(* IEC 61131-3 sources: POMIRTS_lab3/AS/Library_2/ArCert, 3 files *)

(* ---- ArCert.typ ---- *)
 TYPE
	ArCertDetailsType : STRUCT				(*certificate details*)
		Name			: STRING[255]; 			(*certificate name*)
		Issuer			: STRING[255];			(*issuer (CN)*)
		Subject			: STRING[255];			(*subject (CN)*)
		ValidFrom		: DTStructure;			(*valid from date*)
		ValidTo			: DTStructure;			(*valid to date*)
		Version			: DINT;					(*version*)
		SerialNumber	: STRING[39];			(*serial number*)
	END_STRUCT;

	ArCertCRLDetailsType : STRUCT			(*detail information of a certificate revocation list (CRL)*)
		Name			: STRING[255]; 			(*CRL name*)
		Issuer			: STRING[255]; 			(*issuer*)
		EffectiveDate	: DTStructure;			(*effective date*)
		NextUpdate		: DTStructure;			(*next update*)
		Version			: DINT;					(*version*)
		CRLNumber      	: STRING[39]; 			(*CRL number*)
	END_STRUCT;

    ArCertKeySizeEnum :
        (
            arCERT_KEY_SIZE_1024_BITS := 1,		(*encryption with a key with 1024 bits*)
            arCERT_KEY_SIZE_2048_BITS := 2,		(*encryption with a key with 2048 bits*)
            arCERT_KEY_SIZE_4096_BITS := 3		(*encryption with a key with 4096 bits*)
        );

    ArCertAsyncInternalType : STRUCT
        FBStateCtx		: ArFBStateInternalType;
		AsyFuMaCtx		: ArFBAsyFuMaInternalType;
    END_STRUCT;
END_TYPE

(* ---- ArCert.fun ---- *)
{REDUND_CONTEXT} {REDUND_UNREPLICABLE} FUNCTION_BLOCK ArCertImportOwn   				(*imports an existing own certificate from buffer*)
	VAR_INPUT
		Execute			: BOOL; 			(*starts execution*) 			(**) (*#PAR*)
		Name 			: STRING[255];		(*name of the own certificate*) 	(**) (*#PAR*)
		Data			: UDINT; 			(*pointer to certificate data*) (**) (*#PAR*)
		DataSize 		: UDINT;			(*size of certificate data*) 	(**) (*#PAR*)
	END_VAR
	VAR_OUTPUT
		Done			: BOOL;				(*execution done*) 				(**) (*#PAR*)
		Busy			: BOOL;				(*execution running*) 			(**) (*#PAR*)
		Error			: BOOL;				(*execution failed*) 			(**) (*#PAR*)
		StatusID		: DINT;  			(*execution error: see help*) 	(**) (*#PAR*)
	END_VAR
	VAR
		Internal		: ArCertAsyncInternalType;	(*internal variable*)
	END_VAR
END_FUNCTION_BLOCK

{REDUND_CONTEXT} {REDUND_UNREPLICABLE} FUNCTION_BLOCK ArCertExportOwn  				(*exports an own certificate to a buffer*)
	VAR_INPUT
		Execute			: BOOL; 			(*starts execution*) 			(**) (*#PAR*)
		Name 			: STRING[255];		(*name of the own certificate*) 	(**) (*#PAR*)
		Data			: UDINT; 			(*pointer to buffer for exported certificate data*) (**) (*#PAR*)
		DataSize		: UDINT;			(*buffer size*) 				(**) (*#PAR*)
	END_VAR
	VAR_OUTPUT
		Done			: BOOL;				(*execution done*) 				(**) (*#PAR*)
		Busy			: BOOL;				(*execution running*) 			(**) (*#PAR*)
		Error			: BOOL;				(*execution failed*) 			(**) (*#PAR*)
		StatusID		: DINT;  			(*execution error: see help*) 	(**) (*#PAR*)
		NeededDataSize 	: UDINT;			(*needed buffer size*) 				(**) (*#PAR*)
	END_VAR
	VAR
		Internal		: ArCertAsyncInternalType;	(*internal variable*)
	END_VAR
END_FUNCTION_BLOCK

{REDUND_CONTEXT} {REDUND_UNREPLICABLE} FUNCTION_BLOCK ArCertDeleteOwn  				(*deletes an own certificate*)
	VAR_INPUT
		Execute			: BOOL; 			(*starts execution*) 			(**) (*#PAR*)
		Name 			: STRING[255];		(*name of the own certificate*) 	(**) (*#PAR*)
	END_VAR
	VAR_OUTPUT
		Done			: BOOL;				(*execution done*) 				(**) (*#PAR*)
		Busy			: BOOL;				(*execution running*) 			(**) (*#PAR*)
		Error			: BOOL;				(*execution failed*) 			(**) (*#PAR*)
		StatusID		: DINT;  			(*execution error: see help*) 	(**) (*#PAR*)
	END_VAR
	VAR
		Internal		: ArCertAsyncInternalType;	(*internal variable*)
	END_VAR
END_FUNCTION_BLOCK

{REDUND_CONTEXT} {REDUND_UNREPLICABLE} FUNCTION_BLOCK ArCertImportThirdParty   				(*imports an existing third party certificate from buffer*)
	VAR_INPUT
		Execute			: BOOL; 			(*starts execution*) 			(**) (*#PAR*)
		Name 			: STRING[255];		(*name of the third party certificate*) 	(**) (*#PAR*)
		Data			: UDINT; 			(*pointer to certificate data*) (**) (*#PAR*)
		DataSize 		: UDINT;			(*size of certificate data*) 	(**) (*#PAR*)
	END_VAR
	VAR_OUTPUT
		Done			: BOOL;				(*execution done*) 				(**) (*#PAR*)
		Busy			: BOOL;				(*execution running*) 			(**) (*#PAR*)
		Error			: BOOL;				(*execution failed*) 			(**) (*#PAR*)
		StatusID		: DINT;  			(*execution error: see help*) 	(**) (*#PAR*)
	END_VAR
	VAR
		Internal		: ArCertAsyncInternalType;	(*internal variable*)
	END_VAR
END_FUNCTION_BLOCK

{REDUND_CONTEXT} {REDUND_UNREPLICABLE} FUNCTION_BLOCK ArCertExportThirdParty  				(*exports a third party certificate to a buffer*)
	VAR_INPUT
		Execute			: BOOL; 			(*starts execution*) 			(**) (*#PAR*)
		Name 			: STRING[255];		(*name of the third party certificate*) 	(**) (*#PAR*)
		Data			: UDINT; 			(*pointer to buffer for exported certificate data*) (**) (*#PAR*)
		DataSize		: UDINT;			(*buffer size*) 				(**) (*#PAR*)
	END_VAR
	VAR_OUTPUT
		Done			: BOOL;				(*execution done*) 				(**) (*#PAR*)
		Busy			: BOOL;				(*execution running*) 			(**) (*#PAR*)
		Error			: BOOL;				(*execution failed*) 			(**) (*#PAR*)
		StatusID		: DINT;  			(*execution error: see help*) 	(**) (*#PAR*)
		NeededDataSize 	: UDINT;			(*needed buffer size*) 				(**) (*#PAR*)
	END_VAR
	VAR
		Internal		: ArCertAsyncInternalType;	(*internal variable*)
	END_VAR
END_FUNCTION_BLOCK

{REDUND_CONTEXT} {REDUND_UNREPLICABLE} FUNCTION_BLOCK ArCertDeleteThirdParty  				(*deletes a third party certificate*)
	VAR_INPUT
		Execute			: BOOL; 			(*starts execution*) 			(**) (*#PAR*)
		Name 			: STRING[255];		(*name of the third party certificate*) 	(**) (*#PAR*)
	END_VAR
	VAR_OUTPUT
		Done			: BOOL;				(*execution done*) 				(**) (*#PAR*)
		Busy			: BOOL;				(*execution running*) 			(**) (*#PAR*)
		Error			: BOOL;				(*execution failed*) 			(**) (*#PAR*)
		StatusID		: DINT;  			(*execution error: see help*) 	(**) (*#PAR*)
	END_VAR
	VAR
		Internal		: ArCertAsyncInternalType;	(*internal variable*)
	END_VAR
END_FUNCTION_BLOCK

{REDUND_CONTEXT} {REDUND_UNREPLICABLE} FUNCTION_BLOCK ArCertImportPrivateKey		(*imports an existing private key from buffer*)
	VAR_INPUT
		Execute			: BOOL; 			(*starts execution*) 			(**) (*#PAR*)
		Name 			: STRING[255];		(*name of the private key*) 	(**) (*#PAR*)
		Data			: UDINT; 			(*pointer to private key data*) (**) (*#PAR*)
		DataSize 		: UDINT;			(*size of private key data*) 	(**) (*#PAR*)
	END_VAR
	VAR_OUTPUT
		Done			: BOOL;				(*execution done*) 				(**) (*#PAR*)
		Busy			: BOOL;				(*execution running*) 			(**) (*#PAR*)
		Error			: BOOL;				(*execution failed*) 			(**) (*#PAR*)
		StatusID		: DINT;  			(*execution error: see help*) 	(**) (*#PAR*)
	END_VAR
	VAR
		Internal		: ArCertAsyncInternalType;	(*internal variable*)
	END_VAR
END_FUNCTION_BLOCK

{REDUND_CONTEXT} {REDUND_UNREPLICABLE} FUNCTION_BLOCK ArCertExportPrivateKey  		(*exports a private key to a buffer*)
	VAR_INPUT
		Execute			: BOOL; 			(*starts execution*) 			(**) (*#PAR*)
		Name 			: STRING[255];		(*name of the private key*) 	(**) (*#PAR*)
		Data			: UDINT; 			(*pointer to buffer for exported private key data*) (**) (*#PAR*)
		DataSize		: UDINT;			(*buffer size*) 				(**) (*#PAR*)
	END_VAR
	VAR_OUTPUT
		Done			: BOOL;				(*execution done*) 				(**) (*#PAR*)
		Busy			: BOOL;				(*execution running*) 			(**) (*#PAR*)
		Error			: BOOL;				(*execution failed*) 			(**) (*#PAR*)
		StatusID		: DINT;  			(*execution error: see help*) 	(**) (*#PAR*)
		NeededDataSize 	: UDINT;			(*needed buffer size*) 				(**) (*#PAR*)
	END_VAR
	VAR
		Internal		: ArCertAsyncInternalType;	(*internal variable*)
	END_VAR
END_FUNCTION_BLOCK

{REDUND_CONTEXT} {REDUND_UNREPLICABLE} FUNCTION_BLOCK ArCertDeletePrivateKey		(*deletes a private key*)
	VAR_INPUT
		Execute			: BOOL; 			(*starts execution*) 			(**) (*#PAR*)
		Name 			: STRING[255];		(*name of the private key*) 	(**) (*#PAR*)
	END_VAR
	VAR_OUTPUT
		Done			: BOOL;				(*execution done*) 				(**) (*#PAR*)
		Busy			: BOOL;				(*execution running*) 			(**) (*#PAR*)
		Error			: BOOL;				(*execution failed*) 			(**) (*#PAR*)
		StatusID		: DINT;  			(*execution error: see help*) 	(**) (*#PAR*)
	END_VAR
	VAR
		Internal		: ArCertAsyncInternalType;	(*internal variable*)
	END_VAR
END_FUNCTION_BLOCK

{REDUND_CONTEXT} {REDUND_UNREPLICABLE} FUNCTION_BLOCK ArCertImportCRL 				(*imports a certificate revocation list from buffer*)
	VAR_INPUT
		Execute			: BOOL; 			(*starts execution*) 			(**) (*#PAR*)
		Name 			: STRING[255];		(*name of the certificate revocation list*) 	(**) (*#PAR*)
		Data			: UDINT; 			(*pointer to certificate data*) (**) (*#PAR*)
		DataSize 		: UDINT;			(*size of certificate data*) 	(**) (*#PAR*)
	END_VAR
	VAR_OUTPUT
		Done			: BOOL;				(*execution done*) 				(**) (*#PAR*)
		Busy			: BOOL;				(*execution running*) 			(**) (*#PAR*)
		Error			: BOOL;				(*execution failed*) 			(**) (*#PAR*)
		StatusID		: DINT;  			(*execution error: see help*) 	(**) (*#PAR*)
	END_VAR
	VAR
		Internal		: ArCertAsyncInternalType;	(*internal variable*)
	END_VAR
END_FUNCTION_BLOCK

{REDUND_CONTEXT} {REDUND_UNREPLICABLE} FUNCTION_BLOCK ArCertExportCRL 				(*exports a certificate revocation list to a buffer*)
	VAR_INPUT
		Execute			: BOOL; 			(*starts execution*) 			(**) (*#PAR*)
		Name 			: STRING[255];		(*name of the certificate revocation list*) 	(**) (*#PAR*)
		Data			: UDINT; 			(*pointer to buffer for exported CRL data*) (**) (*#PAR*)
		DataSize		: UDINT;			(*buffer size*) 				(**) (*#PAR*)
	END_VAR
	VAR_OUTPUT
		Done			: BOOL;				(*execution done*) 				(**) (*#PAR*)
		Busy			: BOOL;				(*execution running*) 			(**) (*#PAR*)
		Error			: BOOL;				(*execution failed*) 			(**) (*#PAR*)
		StatusID		: DINT;  			(*execution error: see help*) 	(**) (*#PAR*)
		NeededDataSize : UDINT;				(*needed buffer size*) 				(**) (*#PAR*)
	END_VAR
	VAR
		Internal		: ArCertAsyncInternalType;	(*internal variable*)
	END_VAR
END_FUNCTION_BLOCK

{REDUND_CONTEXT} {REDUND_UNREPLICABLE} FUNCTION_BLOCK ArCertDeleteCRL  			(*deletes a certificate revocation list*)
	VAR_INPUT
		Execute			: BOOL; 			(*starts execution*) 			(**) (*#PAR*)
		Name 			: STRING[255];		(*name of the certificate revocation list*) 	(**) (*#PAR*)
	END_VAR
	VAR_OUTPUT
		Done			: BOOL;				(*execution done*) 				(**) (*#PAR*)
		Busy			: BOOL;				(*execution running*) 			(**) (*#PAR*)
		Error			: BOOL;				(*execution failed*) 			(**) (*#PAR*)
		StatusID		: DINT;  			(*execution error: see help*) 	(**) (*#PAR*)
	END_VAR
	VAR
		Internal		: ArCertAsyncInternalType;	(*internal variable*)
	END_VAR
END_FUNCTION_BLOCK

{REDUND_CONTEXT} {REDUND_UNREPLICABLE} FUNCTION_BLOCK ArCertGenerate       		(*generates a self-signed certificate and a private key*)
	VAR_INPUT
		Execute			: BOOL; 			(*starts execution*) 			(**) (*#PAR*)
		Name 			: STRING[255];		(*name of the certificate*) 	(**) (*#PAR*)
		PrivateKeyName 	: STRING[255];		(*name of the private key*) 	(**) (*#PAR*)
		KeySize 		: ArCertKeySizeEnum;(*size of key for certificate generation*) 	(**) (*#PAR*)
		CountryCode		: STRING[9];		(*country code*)		 		(**) (*#PAR*)
		StateProvince	: STRING[513];		(*state*) 						(**) (*#PAR*)
		Locality		: STRING[513];		(*locality*) 					(**) (*#PAR*)
		Organization 	: STRING[255];		(*organization*) 				(**) (*#PAR*)
		OrganizationUnit: STRING[255];		(*organization unit*) 			(**) (*#PAR*)
		ContactEmail 	: STRING[513];		(*contact email*)			 	(**) (*#PAR*)
		CommonName 		: STRING[255];		(*common name*) 				(**) (*#PAR*)
		ValidTimeSeconds : UDINT;			(*valid time in seconds*)		(**) (*#PAR*)
	END_VAR
	VAR_OUTPUT
		Done			: BOOL;				(*execution done*) 				(**) (*#PAR*)
		Busy			: BOOL;				(*execution running*) 			(**) (*#PAR*)
		Error			: BOOL;				(*execution failed*) 			(**) (*#PAR*)
		StatusID		: DINT;  			(*execution error: see help*) 	(**) (*#PAR*)
	END_VAR
	VAR
		Internal		: ArCertAsyncInternalType;	(*internal variable*)
	END_VAR
END_FUNCTION_BLOCK

{REDUND_CONTEXT} {REDUND_UNREPLICABLE} FUNCTION_BLOCK ArCertGenerateOpcUA		(*generates a self-signed certificate and a private key*)
	VAR_INPUT
		Execute			: BOOL; 			(*starts execution*) 			(**) (*#PAR*)
		Name 			: STRING[255];		(*name of the certificate*) 	(**) (*#PAR*)
		PrivateKeyName 	: STRING[255];		(*name of the private key*) 	(**) (*#PAR*)
		PrivateKeyPassword : STRING[255];	(*password of the private key*) (**) (*#PAR*)
		KeySize 		: ArCertKeySizeEnum;(*size of key for certificate generation*) 	(**) (*#PAR*)
		CountryCode		: STRING[9];		(*country code*)		 		(**) (*#PAR*)
		StateProvince	: STRING[513];		(*state*) 						(**) (*#PAR*)
		Locality		: STRING[513];		(*locality*) 					(**) (*#PAR*)
		Organization 	: STRING[255];		(*organization*) 				(**) (*#PAR*)
		OrganizationUnit: STRING[255];		(*organization unit*) 			(**) (*#PAR*)
		ContactEmail 	: STRING[513];		(*contact email*)			 	(**) (*#PAR*)
		CommonName 		: STRING[255];		(*common name*) 				(**) (*#PAR*)
		ValidTimeSeconds : UDINT;			(*valid time in seconds*)		(**) (*#PAR*)
		URI				: STRING[255];		(*URI*) 						(**) (*#PAR*)
	END_VAR
	VAR_OUTPUT
		Done			: BOOL;				(*execution done*) 				(**) (*#PAR*)
		Busy			: BOOL;				(*execution running*) 			(**) (*#PAR*)
		Error			: BOOL;				(*execution failed*) 			(**) (*#PAR*)
		StatusID		: DINT;  			(*execution error: see help*) 	(**) (*#PAR*)
	END_VAR
	VAR
		Internal		: ArCertAsyncInternalType;	(*internal variable*)
	END_VAR
END_FUNCTION_BLOCK

{REDUND_CONTEXT} {REDUND_UNREPLICABLE} FUNCTION_BLOCK ArCertGetOwnDetails   			(*gets details of an own certificate*)
	VAR_INPUT
		Execute			: BOOL; 			(*starts execution*) 			(**) (*#PAR*)
		Name 			: STRING[255];		(*name of the own certificate*) 	(**) (*#PAR*)
		Index			: UDINT;			(*index of the certificate*) (**) (*#PAR*)
	END_VAR
	VAR_OUTPUT
		Done			: BOOL;				(*execution done*) 				(**) (*#PAR*)
		Busy			: BOOL;				(*execution running*) 			(**) (*#PAR*)
		Error			: BOOL;				(*execution failed*) 			(**) (*#PAR*)
		StatusID		: DINT;  			(*execution error: see help*) 	(**) (*#PAR*)
		Details			: ArCertDetailsType;(*certificate details*)
	END_VAR
	VAR
		Internal		: ArCertAsyncInternalType;	(*internal variable*)
	END_VAR
END_FUNCTION_BLOCK

{REDUND_CONTEXT} {REDUND_UNREPLICABLE} FUNCTION_BLOCK ArCertGetThirdPartyDetails   			(*gets details of a third party certificate*)
	VAR_INPUT
		Execute			: BOOL; 			(*starts execution*) 			(**) (*#PAR*)
		Name 			: STRING[255];		(*name of the third party certificate*) 	(**) (*#PAR*)
		Index			: UDINT;			(*index of the certificate*) (**) (*#PAR*)
	END_VAR
	VAR_OUTPUT
		Done			: BOOL;				(*execution done*) 				(**) (*#PAR*)
		Busy			: BOOL;				(*execution running*) 			(**) (*#PAR*)
		Error			: BOOL;				(*execution failed*) 			(**) (*#PAR*)
		StatusID		: DINT;  			(*execution error: see help*) 	(**) (*#PAR*)
		Details			: ArCertDetailsType;(*certificate details*)
	END_VAR
	VAR
		Internal		: ArCertAsyncInternalType;	(*internal variable*)
	END_VAR
END_FUNCTION_BLOCK

{REDUND_CONTEXT} {REDUND_UNREPLICABLE} FUNCTION_BLOCK ArCertGetCRLDetails			(*gets details of a certificate revocation list*)
	VAR_INPUT
		Execute			: BOOL; 			(*starts execution*) 			(**) (*#PAR*)
		Name 			: STRING[255];		(*name of the certificate revocation list*) 	(**) (*#PAR*)
		Index			: UDINT;			(*index of the certificate revocation list*) (**) (*#PAR*)
	END_VAR
	VAR_OUTPUT
		Done			: BOOL;				(*execution done*) 				(**) (*#PAR*)
		Busy			: BOOL;				(*execution running*) 			(**) (*#PAR*)
		Error			: BOOL;				(*execution failed*) 			(**) (*#PAR*)
		StatusID		: DINT;  			(*execution error: see help*) 	(**) (*#PAR*)
		Details			: ArCertCRLDetailsType;	(*certificate revocation list details*)
	END_VAR
	VAR
		Internal		: ArCertAsyncInternalType;	(*internal variable*)
	END_VAR
END_FUNCTION_BLOCK

(* ---- ArCert.var ---- *)
VAR CONSTANT
	arCERT_ERR_CERTIFICATE_NOT_FOUND    : DINT := -1070585796;	(*certificate not found*)
	arCERT_ERR_INTERNAL                 : DINT := -1070585795;	(*internal error*)
	arCERT_ERR_BUFFER_SIZE              : DINT := -1070585794;	(*too small buffer size given*)
	arCERT_ERR_CERTIFICATE_EXISTS       : DINT := -1070585793;	(*certificate already exists*)
	arCERT_ERR_CERT_NAME_TOO_LONG       : DINT := -1070585792;	(*too long certificate name*)
	arCERT_ERR_NAME_INVALID             : DINT := -1070585791;	(*invalid name given*)
	arCERT_ERR_DATA_NULL                : DINT := -1070585790;	(*data pointer NULL*)
	arCERT_ERR_DATA_SIZE_INVALID        : DINT := -1070585789;	(*invalid data size given*)
	arCERT_ERR_PRIVATE_KEY_INVALID      : DINT := -1070585788;	(*invalid private key given*)
	arCERT_ERR_KEY_SIZE_INVALID         : DINT := -1070585787;	(*invalid data size given*)
	arCERT_ERR_COUNTRY_CODE_INVALID     : DINT := -1070585786;	(*invalid data size given*)
	arCERT_ERR_VALID_TIME_INVALID       : DINT := -1070585785;	(*invalid data size given*)
	arCERT_ERR_URI_INVALID              : DINT := -1070585784;	(*invalid URI given*)
END_VAR
